// TIA Portal V20 export
// export: Created 2026-10-19T18:38:13.6336931Z, ExportSetting WithDefaults, DisplayName Totally Integrated Automation Portal, DisplayVersion V20 Update 6, DisplayName TIA Portal Openness, DisplayVersion V20 Update 6, DisplayName TIA Portal Version Control Interface, DisplayVersion V20 Update 6, DisplayName SINAMICS Startdrive Advanced, DisplayVersion V20 SP1, DisplayName SINAMICS Startdrive G130, G150, S120, S150, SINAMICS MV, G220, S200, S210, DisplayVersion V20 SP1, DisplayName SINAMICS Startdrive G110M, G120, G120C, G120D, G120P, G115D, DisplayVersion V20 SP1, DisplayName STEP 7 Professional, DisplayVersion V20 Update 6, DisplayName STEP 7 Safety, DisplayVersion V20 Update 2, DisplayName WinCC Basic/Comfort/Advanced, DisplayVersion V20 Update 6, DisplayName WinCC Unified, DisplayVersion V20 Update 6
DATA_BLOCK "System_VTD_DB_1"   // DB128
{ S7_Optimized_Access := 'TRUE' }
VERSION : 0.1
// stored: AutoNumber true, DBAccessibleFromOPCUA true, InstanceOfName System_UDT, InstanceOfType UDT, IsOnlyStoredInLoadMemory false, IsWriteProtectedInAS false
"System_UDT"
   // VAR
   //    Id : UInt := 1;
   //    CancelOrders : Bool := FALSE;
   //    PauseOrders : Bool := FALSE;
   //    ResumeOrders : Bool := FALSE;
   //    OrderSent : Bool := FALSE;
   //    CurrentOrder : UInt := 0;
   //    NextOrder : UInt := 1;
   //    OrderTable : Array[0..99] of "OrderTable_UDT";
   //    StepTable : Array[0..20] of "OrderTable_UDT";
   //    CarParked_Confirm : Bool := FALSE;
   //    Running { ExternalWritable := 'False'} : Bool := FALSE;
   //    IDLE { ExternalWritable := 'False'} : Bool := TRUE;
   //    Error { ExternalWritable := 'False'} : Bool := FALSE;
   //    State { ExternalWritable := 'False'} : USInt := 0;
   //    ResetError { ExternalWritable := 'False'} : Bool := FALSE;
   //    Ready { ExternalWritable := 'False'} : Bool := TRUE;
   //    Selected { ExternalWritable := 'False'} : Bool := TRUE;
   //    Auto_Man { ExternalWritable := 'False'} : Bool := TRUE;
   //    Paused { ExternalWritable := 'False'} : Bool := FALSE;
   //    Watchdog_TimeOut { ExternalWritable := 'False'} : Struct
   //       VTD { ExternalWritable := 'False'} : Bool;
   //       Pallet_InOut { ExternalWritable := 'False'} : Bool;
   //       Shuttle_InOut { ExternalWritable := 'False'} : Bool;
   //       Level_2 { ExternalWritable := 'False'} : Bool;
   //       Level_3 { ExternalWritable := 'False'} : Bool;
   //       Level_4 { ExternalWritable := 'False'} : Bool;
   //       Level_5 { ExternalWritable := 'False'} : Bool;
   //       Level_6 { ExternalWritable := 'False'} : Bool;
   //    END_STRUCT;
   // END_VAR
BEGIN
   OrderTable[0..99].OrderNo := 0;
   OrderTable[0].StepNo := 256;
   OrderTable[1..99].StepNo := 0;
   OrderTable[0..99].PlaceTime := '';
   OrderTable[0..99].Device := '';
   OrderTable[0..99].Sequence := 0;
   OrderTable[0].Status := 'Error';
   OrderTable[1..99].Status := '';
   OrderTable[0].CompleteTime := '06/10/2022 08:58:15';
   OrderTable[1..99].CompleteTime := '';
   OrderTable[0..99].ErrorID := 0;
   StepTable[1..20].OrderNo := 0;
   StepTable[1..20].StepNo := 0;
   StepTable[1..20].PlaceTime := '';
   StepTable[1..20].Device := '';
   StepTable[1..20].Sequence := 0;
   StepTable[1..20].Status := '';
   StepTable[1..20].CompleteTime := '';
   StepTable[1..20].ErrorID := 0;
END_DATA_BLOCK
